Fanuc KAREL source: kc00013.KL

-- PROVISIONAL review KL for V940-1; original PC SHA256 3dabb6e0b8ed78b567ee729ddf9de5ce019cfcede090bdda4d32e473f01565b7
-- Incomplete behavior may be omitted. Consult companion uncertainty JSON. Do not deploy.
PROGRAM KC00013
%NOLOCKGROUP
BEGIN
  -- V9_ZERO_TABLE_METADATA_HINT layout=0002_ascii; no indexed target words; source/name/runtime held
  -- UNRESOLVED_PC offsets 5-39; opcodes 27,22,22,22,22,22,31
  -- UNRESOLVED_PC offsets 44-48; opcodes 7F
END KC00013
